(* IEC 61131-3 sources: s7-to-codesys/tests/POUs/Scenarios/FB_AlarmDelay_ScenarioTest, 9 files *)

(* ---- FB_AlarmDelay_ScenarioTest.decl.st ---- *)
// AUTO-GENERATED — не редактировать: s7conv gen-tests, сценарии scenarios/FB_AlarmDelay.csv
// Правка — в CSV (scenarios/README.md), затем python -m s7conv build-corpus.
// Назначение: тесты поведения сконвертированного FB_AlarmDelay по сценариям CSV (сценариев: 8, строк: 55):
//             один метод-тест на сценарий, строки — по порядку с моделируемым временем GVL_S7Clock.
//             Ожидаемые значения — из CSV (эталонные модели по описанию логики блока), не из
//             результата конвертации.
// Автор:      s7conv 0.1.0 (сгенерировано)
// Версия:     не указана
// Документ:   scenarios/README.md, docs/methodology.md, раздел «Проверка поведения»
FUNCTION_BLOCK FB_AlarmDelay_ScenarioTest EXTENDS coUnit.FB_TestSuite
VAR
    fbActivateAckClear : FB_AlarmDelay;  // свой экземпляр на сценарий
    xActivateAckClearDone : BOOL;  // сценарий выполнен (выполняется один раз)
    fbClearedBeforeAck : FB_AlarmDelay;  // свой экземпляр на сценарий
    xClearedBeforeAckDone : BOOL;  // сценарий выполнен (выполняется один раз)
    fbChatterSuppressed : FB_AlarmDelay;  // свой экземпляр на сценарий
    xChatterSuppressedDone : BOOL;  // сценарий выполнен (выполняется один раз)
    fbReturnDuringOffDelay : FB_AlarmDelay;  // свой экземпляр на сценарий
    xReturnDuringOffDelayDone : BOOL;  // сценарий выполнен (выполняется один раз)
    fbNewActivationAfterOffDelay : FB_AlarmDelay;  // свой экземпляр на сценарий
    xNewActivationAfterOffDelayDone : BOOL;  // сценарий выполнен (выполняется один раз)
    fbDisabled : FB_AlarmDelay;  // свой экземпляр на сценарий
    xDisabledDone : BOOL;  // сценарий выполнен (выполняется один раз)
    fbAckSameCallAsActivation : FB_AlarmDelay;  // свой экземпляр на сценарий
    xAckSameCallAsActivationDone : BOOL;  // сценарий выполнен (выполняется один раз)
    fbAckHeldDuringActivation : FB_AlarmDelay;  // свой экземпляр на сценарий
    xAckHeldDuringActivationDone : BOOL;  // сценарий выполнен (выполняется один раз)
END_VAR

(* ---- AckHeldDuringActivation.method.impl.st ---- *)
// AUTO-GENERATED — не редактировать: scenarios/FB_AlarmDelay.csv, сценарий AckHeldDuringActivation
coUnit.TEST('AckHeldDuringActivation');
IF NOT xAckHeldDuringActivationDone THEN
    xAckHeldDuringActivationDone := TRUE;
    GVL_S7Clock.xSimulation := TRUE;

    // #1, t = 0 мс — условие; кнопка нажата заранее — фронт ack до появления
    GVL_S7Clock.tSimNow := T#0MS;
    fbAckHeldDuringActivation.condition := TRUE;
    fbAckHeldDuringActivation.enable := TRUE;
    fbAckHeldDuringActivation.ack := TRUE;
    fbAckHeldDuringActivation.onDelay := T#5000MS;
    fbAckHeldDuringActivation.offDelay := T#2000MS;
    fbAckHeldDuringActivation();
    AssertEquals_BOOL(Expected := FALSE,
                      Actual := fbAckHeldDuringActivation.active,
                      Message := 'AckHeldDuringActivation#1 active');
    AssertEquals_BOOL(Expected := FALSE,
                      Actual := fbAckHeldDuringActivation.unacked,
                      Message := 'AckHeldDuringActivation#1 unacked');
    AssertEquals_BOOL(Expected := FALSE,
                      Actual := fbAckHeldDuringActivation.alarm,
                      Message := 'AckHeldDuringActivation#1 alarm');
    AssertEquals_INT(Expected := 0,
                     Actual := fbAckHeldDuringActivation.state,
                     Message := 'AckHeldDuringActivation#1 state');
    AssertEquals_DINT(Expected := 0,
                      Actual := fbAckHeldDuringActivation.count,
                      Message := 'AckHeldDuringActivation#1 count');

    // #2, t = 5200 мс — появление №1 при удерживаемой кнопке: не квитирован
    GVL_S7Clock.tSimNow := T#5200MS;
    fbAckHeldDuringActivation();
    AssertEquals_BOOL(Expected := TRUE,
                      Actual := fbAckHeldDuringActivation.active,
                      Message := 'AckHeldDuringActivation#2 active');
    AssertEquals_BOOL(Expected := TRUE,
                      Actual := fbAckHeldDuringActivation.unacked,
                      Message := 'AckHeldDuringActivation#2 unacked');
    AssertEquals_BOOL(Expected := TRUE,
                      Actual := fbAckHeldDuringActivation.alarm,
                      Message := 'AckHeldDuringActivation#2 alarm');
    AssertEquals_INT(Expected := 1,
                     Actual := fbAckHeldDuringActivation.state,
                     Message := 'AckHeldDuringActivation#2 state');
    AssertEquals_DINT(Expected := 1,
                      Actual := fbAckHeldDuringActivation.count,
                      Message := 'AckHeldDuringActivation#2 count');

    // #3, t = 5400 мс — кнопка всё ещё нажата, фронта нет: не квитирован
    GVL_S7Clock.tSimNow := T#5400MS;
    fbAckHeldDuringActivation();
    AssertEquals_BOOL(Expected := TRUE,
                      Actual := fbAckHeldDuringActivation.active,
                      Message := 'AckHeldDuringActivation#3 active');
    AssertEquals_BOOL(Expected := TRUE,
                      Actual := fbAckHeldDuringActivation.unacked,
                      Message := 'AckHeldDuringActivation#3 unacked');
    AssertEquals_BOOL(Expected := TRUE,
                      Actual := fbAckHeldDuringActivation.alarm,
                      Message := 'AckHeldDuringActivation#3 alarm');
    AssertEquals_INT(Expected := 1,
                     Actual := fbAckHeldDuringActivation.state,
                     Message := 'AckHeldDuringActivation#3 state');
    AssertEquals_DINT(Expected := 1,
                      Actual := fbAckHeldDuringActivation.count,
                      Message := 'AckHeldDuringActivation#3 count');

    // #4, t = 5600 мс — кнопка отпущена
    GVL_S7Clock.tSimNow := T#5600MS;
    fbAckHeldDuringActivation.ack := FALSE;
    fbAckHeldDuringActivation();
    AssertEquals_BOOL(Expected := TRUE,
                      Actual := fbAckHeldDuringActivation.active,
                      Message := 'AckHeldDuringActivation#4 active');
    AssertEquals_BOOL(Expected := TRUE,
                      Actual := fbAckHeldDuringActivation.unacked,
                      Message := 'AckHeldDuringActivation#4 unacked');
    AssertEquals_BOOL(Expected := TRUE,
                      Actual := fbAckHeldDuringActivation.alarm,
                      Message := 'AckHeldDuringActivation#4 alarm');
    AssertEquals_INT(Expected := 1,
                     Actual := fbAckHeldDuringActivation.state,
                     Message := 'AckHeldDuringActivation#4 state');
    AssertEquals_DINT(Expected := 1,
                      Actual := fbAckHeldDuringActivation.count,
                      Message := 'AckHeldDuringActivation#4 count');

    // #5, t = 5800 мс — новый фронт: квитирован
    GVL_S7Clock.tSimNow := T#5800MS;
    fbAckHeldDuringActivation.ack := TRUE;
    fbAckHeldDuringActivation();
    AssertEquals_BOOL(Expected := TRUE,
                      Actual := fbAckHeldDuringActivation.active,
                      Message := 'AckHeldDuringActivation#5 active');
    AssertEquals_BOOL(Expected := FALSE,
                      Actual := fbAckHeldDuringActivation.unacked,
                      Message := 'AckHeldDuringActivation#5 unacked');
    AssertEquals_BOOL(Expected := TRUE,
                      Actual := fbAckHeldDuringActivation.alarm,
                      Message := 'AckHeldDuringActivation#5 alarm');
    AssertEquals_INT(Expected := 2,
                     Actual := fbAckHeldDuringActivation.state,
                     Message := 'AckHeldDuringActivation#5 state');
    AssertEquals_DINT(Expected := 1,
                      Actual := fbAckHeldDuringActivation.count,
                      Message := 'AckHeldDuringActivation#5 count');

    GVL_S7Clock.xSimulation := FALSE;
END_IF
coUnit.TEST_FINISHED();

(* ---- AckSameCallAsActivation.method.impl.st ---- *)
// AUTO-GENERATED — не редактировать: scenarios/FB_AlarmDelay.csv, сценарий AckSameCallAsActivation
coUnit.TEST('AckSameCallAsActivation');
IF NOT xAckSameCallAsActivationDone THEN
    xAckSameCallAsActivationDone := TRUE;
    GVL_S7Clock.xSimulation := TRUE;

    // #1, t = 0 мс — условие
    GVL_S7Clock.tSimNow := T#0MS;
    fbAckSameCallAsActivation.condition := TRUE;
    fbAckSameCallAsActivation.enable := TRUE;
    fbAckSameCallAsActivation.ack := FALSE;
    fbAckSameCallAsActivation.onDelay := T#5000MS;
    fbAckSameCallAsActivation.offDelay := T#2000MS;
    fbAckSameCallAsActivation();
    AssertEquals_BOOL(Expected := FALSE,
                      Actual := fbAckSameCallAsActivation.active,
                      Message := 'AckSameCallAsActivation#1 active');
    AssertEquals_BOOL(Expected := FALSE,
                      Actual := fbAckSameCallAsActivation.unacked,
                      Message := 'AckSameCallAsActivation#1 unacked');
    AssertEquals_BOOL(Expected := FALSE,
                      Actual := fbAckSameCallAsActivation.alarm,
                      Message := 'AckSameCallAsActivation#1 alarm');
    AssertEquals_INT(Expected := 0,
                     Actual := fbAckSameCallAsActivation.state,
                     Message := 'AckSameCallAsActivation#1 state');
    AssertEquals_DINT(Expected := 0,
                      Actual := fbAckSameCallAsActivation.count,
                      Message := 'AckSameCallAsActivation#1 count');

    // #2, t = 5200 мс — появление и фронт ack в одном вызове: не квитирован
    GVL_S7Clock.tSimNow := T#5200MS;
    fbAckSameCallAsActivation.ack := TRUE;
    fbAckSameCallAsActivation();
    AssertEquals_BOOL(Expected := TRUE,
                      Actual := fbAckSameCallAsActivation.active,
                      Message := 'AckSameCallAsActivation#2 active');
    AssertEquals_BOOL(Expected := TRUE,
                      Actual := fbAckSameCallAsActivation.unacked,
                      Message := 'AckSameCallAsActivation#2 unacked');
    AssertEquals_BOOL(Expected := TRUE,
                      Actual := fbAckSameCallAsActivation.alarm,
                      Message := 'AckSameCallAsActivation#2 alarm');
    AssertEquals_INT(Expected := 1,
                     Actual := fbAckSameCallAsActivation.state,
                     Message := 'AckSameCallAsActivation#2 state');
    AssertEquals_DINT(Expected := 1,
                      Actual := fbAckSameCallAsActivation.count,
                      Message := 'AckSameCallAsActivation#2 count');

    // #3, t = 5400 мс — не квитирован
    GVL_S7Clock.tSimNow := T#5400MS;
    fbAckSameCallAsActivation.ack := FALSE;
    fbAckSameCallAsActivation();
    AssertEquals_BOOL(Expected := TRUE,
                      Actual := fbAckSameCallAsActivation.active,
                      Message := 'AckSameCallAsActivation#3 active');
    AssertEquals_BOOL(Expected := TRUE,
                      Actual := fbAckSameCallAsActivation.unacked,
                      Message := 'AckSameCallAsActivation#3 unacked');
    AssertEquals_BOOL(Expected := TRUE,
                      Actual := fbAckSameCallAsActivation.alarm,
                      Message := 'AckSameCallAsActivation#3 alarm');
    AssertEquals_INT(Expected := 1,
                     Actual := fbAckSameCallAsActivation.state,
                     Message := 'AckSameCallAsActivation#3 state');
    AssertEquals_DINT(Expected := 1,
                      Actual := fbAckSameCallAsActivation.count,
                      Message := 'AckSameCallAsActivation#3 count');

    // #4, t = 5600 мс — квитирован
    GVL_S7Clock.tSimNow := T#5600MS;
    fbAckSameCallAsActivation.ack := TRUE;
    fbAckSameCallAsActivation();
    AssertEquals_BOOL(Expected := TRUE,
                      Actual := fbAckSameCallAsActivation.active,
                      Message := 'AckSameCallAsActivation#4 active');
    AssertEquals_BOOL(Expected := FALSE,
                      Actual := fbAckSameCallAsActivation.unacked,
                      Message := 'AckSameCallAsActivation#4 unacked');
    AssertEquals_BOOL(Expected := TRUE,
                      Actual := fbAckSameCallAsActivation.alarm,
                      Message := 'AckSameCallAsActivation#4 alarm');
    AssertEquals_INT(Expected := 2,
                     Actual := fbAckSameCallAsActivation.state,
                     Message := 'AckSameCallAsActivation#4 state');
    AssertEquals_DINT(Expected := 1,
                      Actual := fbAckSameCallAsActivation.count,
                      Message := 'AckSameCallAsActivation#4 count');

    GVL_S7Clock.xSimulation := FALSE;
END_IF
coUnit.TEST_FINISHED();

(* ---- ActivateAckClear.method.impl.st ---- *)
// AUTO-GENERATED — не редактировать: scenarios/FB_AlarmDelay.csv, сценарий ActivateAckClear
coUnit.TEST('ActivateAckClear');
IF NOT xActivateAckClearDone THEN
    xActivateAckClearDone := TRUE;
    GVL_S7Clock.xSimulation := TRUE;

    // #1, t = 0 мс — норма
    GVL_S7Clock.tSimNow := T#0MS;
    fbActivateAckClear.condition := FALSE;
    fbActivateAckClear.enable := TRUE;
    fbActivateAckClear.ack := FALSE;
    fbActivateAckClear.onDelay := T#5000MS;
    fbActivateAckClear.offDelay := T#2000MS;
    fbActivateAckClear();
    AssertEquals_BOOL(Expected := FALSE, Actual := fbActivateAckClear.active, Message := 'ActivateAckClear#1 active');
    AssertEquals_BOOL(Expected := FALSE, Actual := fbActivateAckClear.unacked, Message := 'ActivateAckClear#1 unacked');
    AssertEquals_BOOL(Expected := FALSE, Actual := fbActivateAckClear.alarm, Message := 'ActivateAckClear#1 alarm');
    AssertEquals_INT(Expected := 0, Actual := fbActivateAckClear.state, Message := 'ActivateAckClear#1 state');
    AssertEquals_DINT(Expected := 0, Actual := fbActivateAckClear.count, Message := 'ActivateAckClear#1 count');

    // #2, t = 1000 мс — условие появилось; отсчёт onDelay с 1.0 с
    GVL_S7Clock.tSimNow := T#1000MS;
    fbActivateAckClear.condition := TRUE;
    fbActivateAckClear();
    AssertEquals_BOOL(Expected := FALSE, Actual := fbActivateAckClear.active, Message := 'ActivateAckClear#2 active');
    AssertEquals_BOOL(Expected := FALSE, Actual := fbActivateAckClear.unacked, Message := 'ActivateAckClear#2 unacked');
    AssertEquals_BOOL(Expected := FALSE, Actual := fbActivateAckClear.alarm, Message := 'ActivateAckClear#2 alarm');
    AssertEquals_INT(Expected := 0, Actual := fbActivateAckClear.state, Message := 'ActivateAckClear#2 state');
    AssertEquals_DINT(Expected := 0, Actual := fbActivateAckClear.count, Message := 'ActivateAckClear#2 count');

    // #3, t = 5800 мс — 4.8 с < 5 с: ещё не активен
    GVL_S7Clock.tSimNow := T#5800MS;
    fbActivateAckClear();
    AssertEquals_BOOL(Expected := FALSE, Actual := fbActivateAckClear.active, Message := 'ActivateAckClear#3 active');
    AssertEquals_BOOL(Expected := FALSE, Actual := fbActivateAckClear.unacked, Message := 'ActivateAckClear#3 unacked');
    AssertEquals_BOOL(Expected := FALSE, Actual := fbActivateAckClear.alarm, Message := 'ActivateAckClear#3 alarm');
    AssertEquals_INT(Expected := 0, Actual := fbActivateAckClear.state, Message := 'ActivateAckClear#3 state');
    AssertEquals_DINT(Expected := 0, Actual := fbActivateAckClear.count, Message := 'ActivateAckClear#3 count');

    // #4, t = 6000 мс, на пороге таймера — 5.0 с = onDelay: активен, не квитирован, появление №1
    GVL_S7Clock.tSimNow := T#6000MS;
    fbActivateAckClear();
    AssertEquals_BOOL(Expected := TRUE, Actual := fbActivateAckClear.active, Message := 'ActivateAckClear#4 active');
    AssertEquals_BOOL(Expected := TRUE, Actual := fbActivateAckClear.unacked, Message := 'ActivateAckClear#4 unacked');
    AssertEquals_BOOL(Expected := TRUE, Actual := fbActivateAckClear.alarm, Message := 'ActivateAckClear#4 alarm');
    AssertEquals_INT(Expected := 1, Actual := fbActivateAckClear.state, Message := 'ActivateAckClear#4 state');
    AssertEquals_DINT(Expected := 1, Actual := fbActivateAckClear.count, Message := 'ActivateAckClear#4 count');

    // #5, t = 6200 мс — активен, не квитирован
    GVL_S7Clock.tSimNow := T#6200MS;
    fbActivateAckClear();
    AssertEquals_BOOL(Expected := TRUE, Actual := fbActivateAckClear.active, Message := 'ActivateAckClear#5 active');
    AssertEquals_BOOL(Expected := TRUE, Actual := fbActivateAckClear.unacked, Message := 'ActivateAckClear#5 unacked');
    AssertEquals_BOOL(Expected := TRUE, Actual := fbActivateAckClear.alarm, Message := 'ActivateAckClear#5 alarm');
    AssertEquals_INT(Expected := 1, Actual := fbActivateAckClear.state, Message := 'ActivateAckClear#5 state');
    AssertEquals_DINT(Expected := 1, Actual := fbActivateAckClear.count, Message := 'ActivateAckClear#5 count');

    // #6, t = 7000 мс — квитирование: активен, квитирован
    GVL_S7Clock.tSimNow := T#7000MS;
    fbActivateAckClear.ack := TRUE;
    fbActivateAckClear();
    AssertEquals_BOOL(Expected := TRUE, Actual := fbActivateAckClear.active, Message := 'ActivateAckClear#6 active');
    AssertEquals_BOOL(Expected := FALSE, Actual := fbActivateAckClear.unacked, Message := 'ActivateAckClear#6 unacked');
    AssertEquals_BOOL(Expected := TRUE, Actual := fbActivateAckClear.alarm, Message := 'ActivateAckClear#6 alarm');
    AssertEquals_INT(Expected := 2, Actual := fbActivateAckClear.state, Message := 'ActivateAckClear#6 state');
    AssertEquals_DINT(Expected := 1, Actual := fbActivateAckClear.count, Message := 'ActivateAckClear#6 count');

    // #7, t = 7500 мс — кнопка отпущена
    GVL_S7Clock.tSimNow := T#7500MS;
    fbActivateAckClear.ack := FALSE;
    fbActivateAckClear();
    AssertEquals_BOOL(Expected := TRUE, Actual := fbActivateAckClear.active, Message := 'ActivateAckClear#7 active');
    AssertEquals_BOOL(Expected := FALSE, Actual := fbActivateAckClear.unacked, Message := 'ActivateAckClear#7 unacked');
    AssertEquals_BOOL(Expected := TRUE, Actual := fbActivateAckClear.alarm, Message := 'ActivateAckClear#7 alarm');
    AssertEquals_INT(Expected := 2, Actual := fbActivateAckClear.state, Message := 'ActivateAckClear#7 state');
    AssertEquals_DINT(Expected := 1, Actual := fbActivateAckClear.count, Message := 'ActivateAckClear#7 count');

    // #8, t = 9000 мс — условие пропало; отсчёт offDelay с 9.0 с, сигнал держится
    GVL_S7Clock.tSimNow := T#9000MS;
    fbActivateAckClear.condition := FALSE;
    fbActivateAckClear();
    AssertEquals_BOOL(Expected := TRUE, Actual := fbActivateAckClear.active, Message := 'ActivateAckClear#8 active');
    AssertEquals_BOOL(Expected := FALSE, Actual := fbActivateAckClear.unacked, Message := 'ActivateAckClear#8 unacked');
    AssertEquals_BOOL(Expected := TRUE, Actual := fbActivateAckClear.alarm, Message := 'ActivateAckClear#8 alarm');
    AssertEquals_INT(Expected := 2, Actual := fbActivateAckClear.state, Message := 'ActivateAckClear#8 state');
    AssertEquals_DINT(Expected := 1, Actual := fbActivateAckClear.count, Message := 'ActivateAckClear#8 count');

    // #9, t = 10800 мс — 1.8 с < 2 с: ещё активен
    GVL_S7Clock.tSimNow := T#10800MS;
    fbActivateAckClear();
    AssertEquals_BOOL(Expected := TRUE, Actual := fbActivateAckClear.active, Message := 'ActivateAckClear#9 active');
    AssertEquals_BOOL(Expected := FALSE, Actual := fbActivateAckClear.unacked, Message := 'ActivateAckClear#9 unacked');
    AssertEquals_BOOL(Expected := TRUE, Actual := fbActivateAckClear.alarm, Message := 'ActivateAckClear#9 alarm');
    AssertEquals_INT(Expected := 2, Actual := fbActivateAckClear.state, Message := 'ActivateAckClear#9 state');
    AssertEquals_DINT(Expected := 1, Actual := fbActivateAckClear.count, Message := 'ActivateAckClear#9 count');

    // #10, t = 11000 мс, на пороге таймера — 2.0 с = offDelay: снят, квитирован — норма
    GVL_S7Clock.tSimNow := T#11000MS;
    fbActivateAckClear();
    AssertEquals_BOOL(Expected := FALSE, Actual := fbActivateAckClear.active, Message := 'ActivateAckClear#10 active');
    AssertEquals_BOOL(Expected := FALSE,
                      Actual := fbActivateAckClear.unacked,
                      Message := 'ActivateAckClear#10 unacked');
    AssertEquals_BOOL(Expected := FALSE, Actual := fbActivateAckClear.alarm, Message := 'ActivateAckClear#10 alarm');
    AssertEquals_INT(Expected := 0, Actual := fbActivateAckClear.state, Message := 'ActivateAckClear#10 state');
    AssertEquals_DINT(Expected := 1, Actual := fbActivateAckClear.count, Message := 'ActivateAckClear#10 count');

    // #11, t = 11200 мс — норма
    GVL_S7Clock.tSimNow := T#11200MS;
    fbActivateAckClear();
    AssertEquals_BOOL(Expected := FALSE, Actual := fbActivateAckClear.active, Message := 'ActivateAckClear#11 active');
    AssertEquals_BOOL(Expected := FALSE,
                      Actual := fbActivateAckClear.unacked,
                      Message := 'ActivateAckClear#11 unacked');
    AssertEquals_BOOL(Expected := FALSE, Actual := fbActivateAckClear.alarm, Message := 'ActivateAckClear#11 alarm');
    AssertEquals_INT(Expected := 0, Actual := fbActivateAckClear.state, Message := 'ActivateAckClear#11 state');
    AssertEquals_DINT(Expected := 1, Actual := fbActivateAckClear.count, Message := 'ActivateAckClear#11 count');

    GVL_S7Clock.xSimulation := FALSE;
END_IF
coUnit.TEST_FINISHED();

(* ---- ChatterSuppressed.method.impl.st ---- *)
// AUTO-GENERATED — не редактировать: scenarios/FB_AlarmDelay.csv, сценарий ChatterSuppressed
coUnit.TEST('ChatterSuppressed');
IF NOT xChatterSuppressedDone THEN
    xChatterSuppressedDone := TRUE;
    GVL_S7Clock.xSimulation := TRUE;

    // #1, t = 0 мс — условие
    GVL_S7Clock.tSimNow := T#0MS;
    fbChatterSuppressed.condition := TRUE;
    fbChatterSuppressed.enable := TRUE;
    fbChatterSuppressed.ack := FALSE;
    fbChatterSuppressed.onDelay := T#5000MS;
    fbChatterSuppressed.offDelay := T#2000MS;
    fbChatterSuppressed();
    AssertEquals_BOOL(Expected := FALSE, Actual := fbChatterSuppressed.active, Message := 'ChatterSuppressed#1 active');
    AssertEquals_BOOL(Expected := FALSE,
                      Actual := fbChatterSuppressed.unacked,
                      Message := 'ChatterSuppressed#1 unacked');
    AssertEquals_BOOL(Expected := FALSE, Actual := fbChatterSuppressed.alarm, Message := 'ChatterSuppressed#1 alarm');
    AssertEquals_INT(Expected := 0, Actual := fbChatterSuppressed.state, Message := 'ChatterSuppressed#1 state');
    AssertEquals_DINT(Expected := 0, Actual := fbChatterSuppressed.count, Message := 'ChatterSuppressed#1 count');

    // #2, t = 3000 мс — пропало через 3 с
    GVL_S7Clock.tSimNow := T#3000MS;
    fbChatterSuppressed.condition := FALSE;
    fbChatterSuppressed();
    AssertEquals_BOOL(Expected := FALSE, Actual := fbChatterSuppressed.active, Message := 'ChatterSuppressed#2 active');
    AssertEquals_BOOL(Expected := FALSE,
                      Actual := fbChatterSuppressed.unacked,
                      Message := 'ChatterSuppressed#2 unacked');
    AssertEquals_BOOL(Expected := FALSE, Actual := fbChatterSuppressed.alarm, Message := 'ChatterSuppressed#2 alarm');
    AssertEquals_INT(Expected := 0, Actual := fbChatterSuppressed.state, Message := 'ChatterSuppressed#2 state');
    AssertEquals_DINT(Expected := 0, Actual := fbChatterSuppressed.count, Message := 'ChatterSuppressed#2 count');

    // #3, t = 3500 мс — снова; отсчёт заново с 3.5 с
    GVL_S7Clock.tSimNow := T#3500MS;
    fbChatterSuppressed.condition := TRUE;
    fbChatterSuppressed();
    AssertEquals_BOOL(Expected := FALSE, Actual := fbChatterSuppressed.active, Message := 'ChatterSuppressed#3 active');
    AssertEquals_BOOL(Expected := FALSE,
                      Actual := fbChatterSuppressed.unacked,
                      Message := 'ChatterSuppressed#3 unacked');
    AssertEquals_BOOL(Expected := FALSE, Actual := fbChatterSuppressed.alarm, Message := 'ChatterSuppressed#3 alarm');
    AssertEquals_INT(Expected := 0, Actual := fbChatterSuppressed.state, Message := 'ChatterSuppressed#3 state');
    AssertEquals_DINT(Expected := 0, Actual := fbChatterSuppressed.count, Message := 'ChatterSuppressed#3 count');

    // #4, t = 8000 мс — 4.5 с < 5 с: не активен
    GVL_S7Clock.tSimNow := T#8000MS;
    fbChatterSuppressed();
    AssertEquals_BOOL(Expected := FALSE, Actual := fbChatterSuppressed.active, Message := 'ChatterSuppressed#4 active');
    AssertEquals_BOOL(Expected := FALSE,
                      Actual := fbChatterSuppressed.unacked,
                      Message := 'ChatterSuppressed#4 unacked');
    AssertEquals_BOOL(Expected := FALSE, Actual := fbChatterSuppressed.alarm, Message := 'ChatterSuppressed#4 alarm');
    AssertEquals_INT(Expected := 0, Actual := fbChatterSuppressed.state, Message := 'ChatterSuppressed#4 state');
    AssertEquals_DINT(Expected := 0, Actual := fbChatterSuppressed.count, Message := 'ChatterSuppressed#4 count');

    // #5, t = 8300 мс — пропало
    GVL_S7Clock.tSimNow := T#8300MS;
    fbChatterSuppressed.condition := FALSE;
    fbChatterSuppressed();
    AssertEquals_BOOL(Expected := FALSE, Actual := fbChatterSuppressed.active, Message := 'ChatterSuppressed#5 active');
    AssertEquals_BOOL(Expected := FALSE,
                      Actual := fbChatterSuppressed.unacked,
                      Message := 'ChatterSuppressed#5 unacked');
    AssertEquals_BOOL(Expected := FALSE, Actual := fbChatterSuppressed.alarm, Message := 'ChatterSuppressed#5 alarm');
    AssertEquals_INT(Expected := 0, Actual := fbChatterSuppressed.state, Message := 'ChatterSuppressed#5 state');
    AssertEquals_DINT(Expected := 0, Actual := fbChatterSuppressed.count, Message := 'ChatterSuppressed#5 count');

    // #6, t = 9000 мс — появлений нет
    GVL_S7Clock.tSimNow := T#9000MS;
    fbChatterSuppressed();
    AssertEquals_BOOL(Expected := FALSE, Actual := fbChatterSuppressed.active, Message := 'ChatterSuppressed#6 active');
    AssertEquals_BOOL(Expected := FALSE,
                      Actual := fbChatterSuppressed.unacked,
                      Message := 'ChatterSuppressed#6 unacked');
    AssertEquals_BOOL(Expected := FALSE, Actual := fbChatterSuppressed.alarm, Message := 'ChatterSuppressed#6 alarm');
    AssertEquals_INT(Expected := 0, Actual := fbChatterSuppressed.state, Message := 'ChatterSuppressed#6 state');
    AssertEquals_DINT(Expected := 0, Actual := fbChatterSuppressed.count, Message := 'ChatterSuppressed#6 count');

    GVL_S7Clock.xSimulation := FALSE;
END_IF
coUnit.TEST_FINISHED();

(* ---- ClearedBeforeAck.method.impl.st ---- *)
// AUTO-GENERATED — не редактировать: scenarios/FB_AlarmDelay.csv, сценарий ClearedBeforeAck
coUnit.TEST('ClearedBeforeAck');
IF NOT xClearedBeforeAckDone THEN
    xClearedBeforeAckDone := TRUE;
    GVL_S7Clock.xSimulation := TRUE;

    // #1, t = 0 мс — условие
    GVL_S7Clock.tSimNow := T#0MS;
    fbClearedBeforeAck.condition := TRUE;
    fbClearedBeforeAck.enable := TRUE;
    fbClearedBeforeAck.ack := FALSE;
    fbClearedBeforeAck.onDelay := T#5000MS;
    fbClearedBeforeAck.offDelay := T#2000MS;
    fbClearedBeforeAck();
    AssertEquals_BOOL(Expected := FALSE, Actual := fbClearedBeforeAck.active, Message := 'ClearedBeforeAck#1 active');
    AssertEquals_BOOL(Expected := FALSE, Actual := fbClearedBeforeAck.unacked, Message := 'ClearedBeforeAck#1 unacked');
    AssertEquals_BOOL(Expected := FALSE, Actual := fbClearedBeforeAck.alarm, Message := 'ClearedBeforeAck#1 alarm');
    AssertEquals_INT(Expected := 0, Actual := fbClearedBeforeAck.state, Message := 'ClearedBeforeAck#1 state');
    AssertEquals_DINT(Expected := 0, Actual := fbClearedBeforeAck.count, Message := 'ClearedBeforeAck#1 count');

    // #2, t = 5200 мс — активен, появление №1
    GVL_S7Clock.tSimNow := T#5200MS;
    fbClearedBeforeAck();
    AssertEquals_BOOL(Expected := TRUE, Actual := fbClearedBeforeAck.active, Message := 'ClearedBeforeAck#2 active');
    AssertEquals_BOOL(Expected := TRUE, Actual := fbClearedBeforeAck.unacked, Message := 'ClearedBeforeAck#2 unacked');
    AssertEquals_BOOL(Expected := TRUE, Actual := fbClearedBeforeAck.alarm, Message := 'ClearedBeforeAck#2 alarm');
    AssertEquals_INT(Expected := 1, Actual := fbClearedBeforeAck.state, Message := 'ClearedBeforeAck#2 state');
    AssertEquals_DINT(Expected := 1, Actual := fbClearedBeforeAck.count, Message := 'ClearedBeforeAck#2 count');

    // #3, t = 6000 мс — условие пропало
    GVL_S7Clock.tSimNow := T#6000MS;
    fbClearedBeforeAck.condition := FALSE;
    fbClearedBeforeAck();
    AssertEquals_BOOL(Expected := TRUE, Actual := fbClearedBeforeAck.active, Message := 'ClearedBeforeAck#3 active');
    AssertEquals_BOOL(Expected := TRUE, Actual := fbClearedBeforeAck.unacked, Message := 'ClearedBeforeAck#3 unacked');
    AssertEquals_BOOL(Expected := TRUE, Actual := fbClearedBeforeAck.alarm, Message := 'ClearedBeforeAck#3 alarm');
    AssertEquals_INT(Expected := 1, Actual := fbClearedBeforeAck.state, Message := 'ClearedBeforeAck#3 state');
    AssertEquals_DINT(Expected := 1, Actual := fbClearedBeforeAck.count, Message := 'ClearedBeforeAck#3 count');

    // #4, t = 8200 мс — через 2.2 с снят, но не квитирован: состояние 3, индикация есть
    GVL_S7Clock.tSimNow := T#8200MS;
    fbClearedBeforeAck();
    AssertEquals_BOOL(Expected := FALSE, Actual := fbClearedBeforeAck.active, Message := 'ClearedBeforeAck#4 active');
    AssertEquals_BOOL(Expected := TRUE, Actual := fbClearedBeforeAck.unacked, Message := 'ClearedBeforeAck#4 unacked');
    AssertEquals_BOOL(Expected := TRUE, Actual := fbClearedBeforeAck.alarm, Message := 'ClearedBeforeAck#4 alarm');
    AssertEquals_INT(Expected := 3, Actual := fbClearedBeforeAck.state, Message := 'ClearedBeforeAck#4 state');
    AssertEquals_DINT(Expected := 1, Actual := fbClearedBeforeAck.count, Message := 'ClearedBeforeAck#4 count');

    // #5, t = 9000 мс — квитирование: норма
    GVL_S7Clock.tSimNow := T#9000MS;
    fbClearedBeforeAck.ack := TRUE;
    fbClearedBeforeAck();
    AssertEquals_BOOL(Expected := FALSE, Actual := fbClearedBeforeAck.active, Message := 'ClearedBeforeAck#5 active');
    AssertEquals_BOOL(Expected := FALSE, Actual := fbClearedBeforeAck.unacked, Message := 'ClearedBeforeAck#5 unacked');
    AssertEquals_BOOL(Expected := FALSE, Actual := fbClearedBeforeAck.alarm, Message := 'ClearedBeforeAck#5 alarm');
    AssertEquals_INT(Expected := 0, Actual := fbClearedBeforeAck.state, Message := 'ClearedBeforeAck#5 state');
    AssertEquals_DINT(Expected := 1, Actual := fbClearedBeforeAck.count, Message := 'ClearedBeforeAck#5 count');

    // #6, t = 9500 мс — норма
    GVL_S7Clock.tSimNow := T#9500MS;
    fbClearedBeforeAck.ack := FALSE;
    fbClearedBeforeAck();
    AssertEquals_BOOL(Expected := FALSE, Actual := fbClearedBeforeAck.active, Message := 'ClearedBeforeAck#6 active');
    AssertEquals_BOOL(Expected := FALSE, Actual := fbClearedBeforeAck.unacked, Message := 'ClearedBeforeAck#6 unacked');
    AssertEquals_BOOL(Expected := FALSE, Actual := fbClearedBeforeAck.alarm, Message := 'ClearedBeforeAck#6 alarm');
    AssertEquals_INT(Expected := 0, Actual := fbClearedBeforeAck.state, Message := 'ClearedBeforeAck#6 state');
    AssertEquals_DINT(Expected := 1, Actual := fbClearedBeforeAck.count, Message := 'ClearedBeforeAck#6 count');

    GVL_S7Clock.xSimulation := FALSE;
END_IF
coUnit.TEST_FINISHED();

(* ---- Disabled.method.impl.st ---- *)
// AUTO-GENERATED — не редактировать: scenarios/FB_AlarmDelay.csv, сценарий Disabled
coUnit.TEST('Disabled');
IF NOT xDisabledDone THEN
    xDisabledDone := TRUE;
    GVL_S7Clock.xSimulation := TRUE;

    // #1, t = 0 мс — условие
    GVL_S7Clock.tSimNow := T#0MS;
    fbDisabled.condition := TRUE;
    fbDisabled.enable := TRUE;
    fbDisabled.ack := FALSE;
    fbDisabled.onDelay := T#5000MS;
    fbDisabled.offDelay := T#2000MS;
    fbDisabled();
    AssertEquals_BOOL(Expected := FALSE, Actual := fbDisabled.active, Message := 'Disabled#1 active');
    AssertEquals_BOOL(Expected := FALSE, Actual := fbDisabled.unacked, Message := 'Disabled#1 unacked');
    AssertEquals_BOOL(Expected := FALSE, Actual := fbDisabled.alarm, Message := 'Disabled#1 alarm');
    AssertEquals_INT(Expected := 0, Actual := fbDisabled.state, Message := 'Disabled#1 state');
    AssertEquals_DINT(Expected := 0, Actual := fbDisabled.count, Message := 'Disabled#1 count');

    // #2, t = 5200 мс — активен, появление №1
    GVL_S7Clock.tSimNow := T#5200MS;
    fbDisabled();
    AssertEquals_BOOL(Expected := TRUE, Actual := fbDisabled.active, Message := 'Disabled#2 active');
    AssertEquals_BOOL(Expected := TRUE, Actual := fbDisabled.unacked, Message := 'Disabled#2 unacked');
    AssertEquals_BOOL(Expected := TRUE, Actual := fbDisabled.alarm, Message := 'Disabled#2 alarm');
    AssertEquals_INT(Expected := 1, Actual := fbDisabled.state, Message := 'Disabled#2 state');
    AssertEquals_DINT(Expected := 1, Actual := fbDisabled.count, Message := 'Disabled#2 count');

    // #3, t = 6000 мс — выведен из работы: active и unacked сброшены сразу
    GVL_S7Clock.tSimNow := T#6000MS;
    fbDisabled.enable := FALSE;
    fbDisabled();
    AssertEquals_BOOL(Expected := FALSE, Actual := fbDisabled.active, Message := 'Disabled#3 active');
    AssertEquals_BOOL(Expected := FALSE, Actual := fbDisabled.unacked, Message := 'Disabled#3 unacked');
    AssertEquals_BOOL(Expected := FALSE, Actual := fbDisabled.alarm, Message := 'Disabled#3 alarm');
    AssertEquals_INT(Expected := 0, Actual := fbDisabled.state, Message := 'Disabled#3 state');
    AssertEquals_DINT(Expected := 1, Actual := fbDisabled.count, Message := 'Disabled#3 count');

    // #4, t = 7000 мс — выведен
    GVL_S7Clock.tSimNow := T#7000MS;
    fbDisabled();
    AssertEquals_BOOL(Expected := FALSE, Actual := fbDisabled.active, Message := 'Disabled#4 active');
    AssertEquals_BOOL(Expected := FALSE, Actual := fbDisabled.unacked, Message := 'Disabled#4 unacked');
    AssertEquals_BOOL(Expected := FALSE, Actual := fbDisabled.alarm, Message := 'Disabled#4 alarm');
    AssertEquals_INT(Expected := 0, Actual := fbDisabled.state, Message := 'Disabled#4 state');
    AssertEquals_DINT(Expected := 1, Actual := fbDisabled.count, Message := 'Disabled#4 count');

    // #5, t = 8500 мс — выведен (задержка снятия внутри уже истекла)
    GVL_S7Clock.tSimNow := T#8500MS;
    fbDisabled();
    AssertEquals_BOOL(Expected := FALSE, Actual := fbDisabled.active, Message := 'Disabled#5 active');
    AssertEquals_BOOL(Expected := FALSE, Actual := fbDisabled.unacked, Message := 'Disabled#5 unacked');
    AssertEquals_BOOL(Expected := FALSE, Actual := fbDisabled.alarm, Message := 'Disabled#5 alarm');
    AssertEquals_INT(Expected := 0, Actual := fbDisabled.state, Message := 'Disabled#5 state');
    AssertEquals_DINT(Expected := 1, Actual := fbDisabled.count, Message := 'Disabled#5 count');

    // #6, t = 9000 мс — введён: условие есть, onDelay с 9.0 с
    GVL_S7Clock.tSimNow := T#9000MS;
    fbDisabled.enable := TRUE;
    fbDisabled();
    AssertEquals_BOOL(Expected := FALSE, Actual := fbDisabled.active, Message := 'Disabled#6 active');
    AssertEquals_BOOL(Expected := FALSE, Actual := fbDisabled.unacked, Message := 'Disabled#6 unacked');
    AssertEquals_BOOL(Expected := FALSE, Actual := fbDisabled.alarm, Message := 'Disabled#6 alarm');
    AssertEquals_INT(Expected := 0, Actual := fbDisabled.state, Message := 'Disabled#6 state');
    AssertEquals_DINT(Expected := 1, Actual := fbDisabled.count, Message := 'Disabled#6 count');

    // #7, t = 14200 мс — 5.2 с: активен, появление №2
    GVL_S7Clock.tSimNow := T#14200MS;
    fbDisabled();
    AssertEquals_BOOL(Expected := TRUE, Actual := fbDisabled.active, Message := 'Disabled#7 active');
    AssertEquals_BOOL(Expected := TRUE, Actual := fbDisabled.unacked, Message := 'Disabled#7 unacked');
    AssertEquals_BOOL(Expected := TRUE, Actual := fbDisabled.alarm, Message := 'Disabled#7 alarm');
    AssertEquals_INT(Expected := 1, Actual := fbDisabled.state, Message := 'Disabled#7 state');
    AssertEquals_DINT(Expected := 2, Actual := fbDisabled.count, Message := 'Disabled#7 count');

    GVL_S7Clock.xSimulation := FALSE;
END_IF
coUnit.TEST_FINISHED();

(* ---- NewActivationAfterOffDelay.method.impl.st ---- *)
// AUTO-GENERATED — не редактировать: scenarios/FB_AlarmDelay.csv, сценарий NewActivationAfterOffDelay
coUnit.TEST('NewActivationAfterOffDelay');
IF NOT xNewActivationAfterOffDelayDone THEN
    xNewActivationAfterOffDelayDone := TRUE;
    GVL_S7Clock.xSimulation := TRUE;

    // #1, t = 0 мс — условие
    GVL_S7Clock.tSimNow := T#0MS;
    fbNewActivationAfterOffDelay.condition := TRUE;
    fbNewActivationAfterOffDelay.enable := TRUE;
    fbNewActivationAfterOffDelay.ack := FALSE;
    fbNewActivationAfterOffDelay.onDelay := T#5000MS;
    fbNewActivationAfterOffDelay.offDelay := T#2000MS;
    fbNewActivationAfterOffDelay();
    AssertEquals_BOOL(Expected := FALSE,
                      Actual := fbNewActivationAfterOffDelay.active,
                      Message := 'NewActivationAfterOffDelay#1 active');
    AssertEquals_BOOL(Expected := FALSE,
                      Actual := fbNewActivationAfterOffDelay.unacked,
                      Message := 'NewActivationAfterOffDelay#1 unacked');
    AssertEquals_BOOL(Expected := FALSE,
                      Actual := fbNewActivationAfterOffDelay.alarm,
                      Message := 'NewActivationAfterOffDelay#1 alarm');
    AssertEquals_INT(Expected := 0,
                     Actual := fbNewActivationAfterOffDelay.state,
                     Message := 'NewActivationAfterOffDelay#1 state');
    AssertEquals_DINT(Expected := 0,
                      Actual := fbNewActivationAfterOffDelay.count,
                      Message := 'NewActivationAfterOffDelay#1 count');

    // #2, t = 5200 мс — активен, появление №1
    GVL_S7Clock.tSimNow := T#5200MS;
    fbNewActivationAfterOffDelay();
    AssertEquals_BOOL(Expected := TRUE,
                      Actual := fbNewActivationAfterOffDelay.active,
                      Message := 'NewActivationAfterOffDelay#2 active');
    AssertEquals_BOOL(Expected := TRUE,
                      Actual := fbNewActivationAfterOffDelay.unacked,
                      Message := 'NewActivationAfterOffDelay#2 unacked');
    AssertEquals_BOOL(Expected := TRUE,
                      Actual := fbNewActivationAfterOffDelay.alarm,
                      Message := 'NewActivationAfterOffDelay#2 alarm');
    AssertEquals_INT(Expected := 1,
                     Actual := fbNewActivationAfterOffDelay.state,
                     Message := 'NewActivationAfterOffDelay#2 state');
    AssertEquals_DINT(Expected := 1,
                      Actual := fbNewActivationAfterOffDelay.count,
                      Message := 'NewActivationAfterOffDelay#2 count');

    // #3, t = 6000 мс — условие пропало
    GVL_S7Clock.tSimNow := T#6000MS;
    fbNewActivationAfterOffDelay.condition := FALSE;
    fbNewActivationAfterOffDelay();
    AssertEquals_BOOL(Expected := TRUE,
                      Actual := fbNewActivationAfterOffDelay.active,
                      Message := 'NewActivationAfterOffDelay#3 active');
    AssertEquals_BOOL(Expected := TRUE,
                      Actual := fbNewActivationAfterOffDelay.unacked,
                      Message := 'NewActivationAfterOffDelay#3 unacked');
    AssertEquals_BOOL(Expected := TRUE,
                      Actual := fbNewActivationAfterOffDelay.alarm,
                      Message := 'NewActivationAfterOffDelay#3 alarm');
    AssertEquals_INT(Expected := 1,
                     Actual := fbNewActivationAfterOffDelay.state,
                     Message := 'NewActivationAfterOffDelay#3 state');
    AssertEquals_DINT(Expected := 1,
                      Actual := fbNewActivationAfterOffDelay.count,
                      Message := 'NewActivationAfterOffDelay#3 count');

    // #4, t = 7000 мс — вернулось; onDelay с 7.0 с, offDelay ещё идёт
    GVL_S7Clock.tSimNow := T#7000MS;
    fbNewActivationAfterOffDelay.condition := TRUE;
    fbNewActivationAfterOffDelay();
    AssertEquals_BOOL(Expected := TRUE,
                      Actual := fbNewActivationAfterOffDelay.active,
                      Message := 'NewActivationAfterOffDelay#4 active');
    AssertEquals_BOOL(Expected := TRUE,
                      Actual := fbNewActivationAfterOffDelay.unacked,
                      Message := 'NewActivationAfterOffDelay#4 unacked');
    AssertEquals_BOOL(Expected := TRUE,
                      Actual := fbNewActivationAfterOffDelay.alarm,
                      Message := 'NewActivationAfterOffDelay#4 alarm');
    AssertEquals_INT(Expected := 1,
                     Actual := fbNewActivationAfterOffDelay.state,
                     Message := 'NewActivationAfterOffDelay#4 state');
    AssertEquals_DINT(Expected := 1,
                      Actual := fbNewActivationAfterOffDelay.count,
                      Message := 'NewActivationAfterOffDelay#4 count');

    // #5, t = 8200 мс — offDelay 2.2 с истёк: снят, не квитирован — состояние 3
    GVL_S7Clock.tSimNow := T#8200MS;
    fbNewActivationAfterOffDelay();
    AssertEquals_BOOL(Expected := FALSE,
                      Actual := fbNewActivationAfterOffDelay.active,
                      Message := 'NewActivationAfterOffDelay#5 active');
    AssertEquals_BOOL(Expected := TRUE,
                      Actual := fbNewActivationAfterOffDelay.unacked,
                      Message := 'NewActivationAfterOffDelay#5 unacked');
    AssertEquals_BOOL(Expected := TRUE,
                      Actual := fbNewActivationAfterOffDelay.alarm,
                      Message := 'NewActivationAfterOffDelay#5 alarm');
    AssertEquals_INT(Expected := 3,
                     Actual := fbNewActivationAfterOffDelay.state,
                     Message := 'NewActivationAfterOffDelay#5 state');
    AssertEquals_DINT(Expected := 1,
                      Actual := fbNewActivationAfterOffDelay.count,
                      Message := 'NewActivationAfterOffDelay#5 count');

    // #6, t = 12200 мс — onDelay 5.2 с: активен снова, появление №2
    GVL_S7Clock.tSimNow := T#12200MS;
    fbNewActivationAfterOffDelay();
    AssertEquals_BOOL(Expected := TRUE,
                      Actual := fbNewActivationAfterOffDelay.active,
                      Message := 'NewActivationAfterOffDelay#6 active');
    AssertEquals_BOOL(Expected := TRUE,
                      Actual := fbNewActivationAfterOffDelay.unacked,
                      Message := 'NewActivationAfterOffDelay#6 unacked');
    AssertEquals_BOOL(Expected := TRUE,
                      Actual := fbNewActivationAfterOffDelay.alarm,
                      Message := 'NewActivationAfterOffDelay#6 alarm');
    AssertEquals_INT(Expected := 1,
                     Actual := fbNewActivationAfterOffDelay.state,
                     Message := 'NewActivationAfterOffDelay#6 state');
    AssertEquals_DINT(Expected := 2,
                      Actual := fbNewActivationAfterOffDelay.count,
                      Message := 'NewActivationAfterOffDelay#6 count');

    // #7, t = 13000 мс — квитирование
    GVL_S7Clock.tSimNow := T#13000MS;
    fbNewActivationAfterOffDelay.ack := TRUE;
    fbNewActivationAfterOffDelay();
    AssertEquals_BOOL(Expected := TRUE,
                      Actual := fbNewActivationAfterOffDelay.active,
                      Message := 'NewActivationAfterOffDelay#7 active');
    AssertEquals_BOOL(Expected := FALSE,
                      Actual := fbNewActivationAfterOffDelay.unacked,
                      Message := 'NewActivationAfterOffDelay#7 unacked');
    AssertEquals_BOOL(Expected := TRUE,
                      Actual := fbNewActivationAfterOffDelay.alarm,
                      Message := 'NewActivationAfterOffDelay#7 alarm');
    AssertEquals_INT(Expected := 2,
                     Actual := fbNewActivationAfterOffDelay.state,
                     Message := 'NewActivationAfterOffDelay#7 state');
    AssertEquals_DINT(Expected := 2,
                      Actual := fbNewActivationAfterOffDelay.count,
                      Message := 'NewActivationAfterOffDelay#7 count');

    GVL_S7Clock.xSimulation := FALSE;
END_IF
coUnit.TEST_FINISHED();

(* ---- ReturnDuringOffDelay.method.impl.st ---- *)
// AUTO-GENERATED — не редактировать: scenarios/FB_AlarmDelay.csv, сценарий ReturnDuringOffDelay
coUnit.TEST('ReturnDuringOffDelay');
IF NOT xReturnDuringOffDelayDone THEN
    xReturnDuringOffDelayDone := TRUE;
    GVL_S7Clock.xSimulation := TRUE;

    // #1, t = 0 мс — условие, offDelay 6 с
    GVL_S7Clock.tSimNow := T#0MS;
    fbReturnDuringOffDelay.condition := TRUE;
    fbReturnDuringOffDelay.enable := TRUE;
    fbReturnDuringOffDelay.ack := FALSE;
    fbReturnDuringOffDelay.onDelay := T#5000MS;
    fbReturnDuringOffDelay.offDelay := T#6000MS;
    fbReturnDuringOffDelay();
    AssertEquals_BOOL(Expected := FALSE,
                      Actual := fbReturnDuringOffDelay.active,
                      Message := 'ReturnDuringOffDelay#1 active');
    AssertEquals_BOOL(Expected := FALSE,
                      Actual := fbReturnDuringOffDelay.unacked,
                      Message := 'ReturnDuringOffDelay#1 unacked');
    AssertEquals_BOOL(Expected := FALSE,
                      Actual := fbReturnDuringOffDelay.alarm,
                      Message := 'ReturnDuringOffDelay#1 alarm');
    AssertEquals_INT(Expected := 0, Actual := fbReturnDuringOffDelay.state, Message := 'ReturnDuringOffDelay#1 state');
    AssertEquals_DINT(Expected := 0, Actual := fbReturnDuringOffDelay.count, Message := 'ReturnDuringOffDelay#1 count');

    // #2, t = 5200 мс — активен, появление №1
    GVL_S7Clock.tSimNow := T#5200MS;
    fbReturnDuringOffDelay();
    AssertEquals_BOOL(Expected := TRUE,
                      Actual := fbReturnDuringOffDelay.active,
                      Message := 'ReturnDuringOffDelay#2 active');
    AssertEquals_BOOL(Expected := TRUE,
                      Actual := fbReturnDuringOffDelay.unacked,
                      Message := 'ReturnDuringOffDelay#2 unacked');
    AssertEquals_BOOL(Expected := TRUE,
                      Actual := fbReturnDuringOffDelay.alarm,
                      Message := 'ReturnDuringOffDelay#2 alarm');
    AssertEquals_INT(Expected := 1, Actual := fbReturnDuringOffDelay.state, Message := 'ReturnDuringOffDelay#2 state');
    AssertEquals_DINT(Expected := 1, Actual := fbReturnDuringOffDelay.count, Message := 'ReturnDuringOffDelay#2 count');

    // #3, t = 5500 мс — квитирован
    GVL_S7Clock.tSimNow := T#5500MS;
    fbReturnDuringOffDelay.ack := TRUE;
    fbReturnDuringOffDelay();
    AssertEquals_BOOL(Expected := TRUE,
                      Actual := fbReturnDuringOffDelay.active,
                      Message := 'ReturnDuringOffDelay#3 active');
    AssertEquals_BOOL(Expected := FALSE,
                      Actual := fbReturnDuringOffDelay.unacked,
                      Message := 'ReturnDuringOffDelay#3 unacked');
    AssertEquals_BOOL(Expected := TRUE,
                      Actual := fbReturnDuringOffDelay.alarm,
                      Message := 'ReturnDuringOffDelay#3 alarm');
    AssertEquals_INT(Expected := 2, Actual := fbReturnDuringOffDelay.state, Message := 'ReturnDuringOffDelay#3 state');
    AssertEquals_DINT(Expected := 1, Actual := fbReturnDuringOffDelay.count, Message := 'ReturnDuringOffDelay#3 count');

    // #4, t = 6000 мс — условие пропало; offDelay с 6.0 с
    GVL_S7Clock.tSimNow := T#6000MS;
    fbReturnDuringOffDelay.condition := FALSE;
    fbReturnDuringOffDelay.ack := FALSE;
    fbReturnDuringOffDelay();
    AssertEquals_BOOL(Expected := TRUE,
                      Actual := fbReturnDuringOffDelay.active,
                      Message := 'ReturnDuringOffDelay#4 active');
    AssertEquals_BOOL(Expected := FALSE,
                      Actual := fbReturnDuringOffDelay.unacked,
                      Message := 'ReturnDuringOffDelay#4 unacked');
    AssertEquals_BOOL(Expected := TRUE,
                      Actual := fbReturnDuringOffDelay.alarm,
                      Message := 'ReturnDuringOffDelay#4 alarm');
    AssertEquals_INT(Expected := 2, Actual := fbReturnDuringOffDelay.state, Message := 'ReturnDuringOffDelay#4 state');
    AssertEquals_DINT(Expected := 1, Actual := fbReturnDuringOffDelay.count, Message := 'ReturnDuringOffDelay#4 count');

    // #5, t = 7000 мс — условие вернулось; onDelay заново с 7.0 с
    GVL_S7Clock.tSimNow := T#7000MS;
    fbReturnDuringOffDelay.condition := TRUE;
    fbReturnDuringOffDelay();
    AssertEquals_BOOL(Expected := TRUE,
                      Actual := fbReturnDuringOffDelay.active,
                      Message := 'ReturnDuringOffDelay#5 active');
    AssertEquals_BOOL(Expected := FALSE,
                      Actual := fbReturnDuringOffDelay.unacked,
                      Message := 'ReturnDuringOffDelay#5 unacked');
    AssertEquals_BOOL(Expected := TRUE,
                      Actual := fbReturnDuringOffDelay.alarm,
                      Message := 'ReturnDuringOffDelay#5 alarm');
    AssertEquals_INT(Expected := 2, Actual := fbReturnDuringOffDelay.state, Message := 'ReturnDuringOffDelay#5 state');
    AssertEquals_DINT(Expected := 1, Actual := fbReturnDuringOffDelay.count, Message := 'ReturnDuringOffDelay#5 count');

    // #6, t = 11800 мс — onDelay 4.8 с, offDelay 5.8 с: ещё активен по задержке снятия
    GVL_S7Clock.tSimNow := T#11800MS;
    fbReturnDuringOffDelay();
    AssertEquals_BOOL(Expected := TRUE,
                      Actual := fbReturnDuringOffDelay.active,
                      Message := 'ReturnDuringOffDelay#6 active');
    AssertEquals_BOOL(Expected := FALSE,
                      Actual := fbReturnDuringOffDelay.unacked,
                      Message := 'ReturnDuringOffDelay#6 unacked');
    AssertEquals_BOOL(Expected := TRUE,
                      Actual := fbReturnDuringOffDelay.alarm,
                      Message := 'ReturnDuringOffDelay#6 alarm');
    AssertEquals_INT(Expected := 2, Actual := fbReturnDuringOffDelay.state, Message := 'ReturnDuringOffDelay#6 state');
    AssertEquals_DINT(Expected := 1, Actual := fbReturnDuringOffDelay.count, Message := 'ReturnDuringOffDelay#6 count');

    // #7, t = 12200 мс — onDelay истёк раньше offDelay: активен без перерыва, счёт не растёт
    GVL_S7Clock.tSimNow := T#12200MS;
    fbReturnDuringOffDelay();
    AssertEquals_BOOL(Expected := TRUE,
                      Actual := fbReturnDuringOffDelay.active,
                      Message := 'ReturnDuringOffDelay#7 active');
    AssertEquals_BOOL(Expected := FALSE,
                      Actual := fbReturnDuringOffDelay.unacked,
                      Message := 'ReturnDuringOffDelay#7 unacked');
    AssertEquals_BOOL(Expected := TRUE,
                      Actual := fbReturnDuringOffDelay.alarm,
                      Message := 'ReturnDuringOffDelay#7 alarm');
    AssertEquals_INT(Expected := 2, Actual := fbReturnDuringOffDelay.state, Message := 'ReturnDuringOffDelay#7 state');
    AssertEquals_DINT(Expected := 1, Actual := fbReturnDuringOffDelay.count, Message := 'ReturnDuringOffDelay#7 count');

    // #8, t = 13000 мс — условие пропало; offDelay с 13.0 с
    GVL_S7Clock.tSimNow := T#13000MS;
    fbReturnDuringOffDelay.condition := FALSE;
    fbReturnDuringOffDelay();
    AssertEquals_BOOL(Expected := TRUE,
                      Actual := fbReturnDuringOffDelay.active,
                      Message := 'ReturnDuringOffDelay#8 active');
    AssertEquals_BOOL(Expected := FALSE,
                      Actual := fbReturnDuringOffDelay.unacked,
                      Message := 'ReturnDuringOffDelay#8 unacked');
    AssertEquals_BOOL(Expected := TRUE,
                      Actual := fbReturnDuringOffDelay.alarm,
                      Message := 'ReturnDuringOffDelay#8 alarm');
    AssertEquals_INT(Expected := 2, Actual := fbReturnDuringOffDelay.state, Message := 'ReturnDuringOffDelay#8 state');
    AssertEquals_DINT(Expected := 1, Actual := fbReturnDuringOffDelay.count, Message := 'ReturnDuringOffDelay#8 count');

    // #9, t = 19200 мс — 6.2 с: снят — норма
    GVL_S7Clock.tSimNow := T#19200MS;
    fbReturnDuringOffDelay();
    AssertEquals_BOOL(Expected := FALSE,
                      Actual := fbReturnDuringOffDelay.active,
                      Message := 'ReturnDuringOffDelay#9 active');
    AssertEquals_BOOL(Expected := FALSE,
                      Actual := fbReturnDuringOffDelay.unacked,
                      Message := 'ReturnDuringOffDelay#9 unacked');
    AssertEquals_BOOL(Expected := FALSE,
                      Actual := fbReturnDuringOffDelay.alarm,
                      Message := 'ReturnDuringOffDelay#9 alarm');
    AssertEquals_INT(Expected := 0, Actual := fbReturnDuringOffDelay.state, Message := 'ReturnDuringOffDelay#9 state');
    AssertEquals_DINT(Expected := 1, Actual := fbReturnDuringOffDelay.count, Message := 'ReturnDuringOffDelay#9 count');

    GVL_S7Clock.xSimulation := FALSE;
END_IF
coUnit.TEST_FINISHED();
